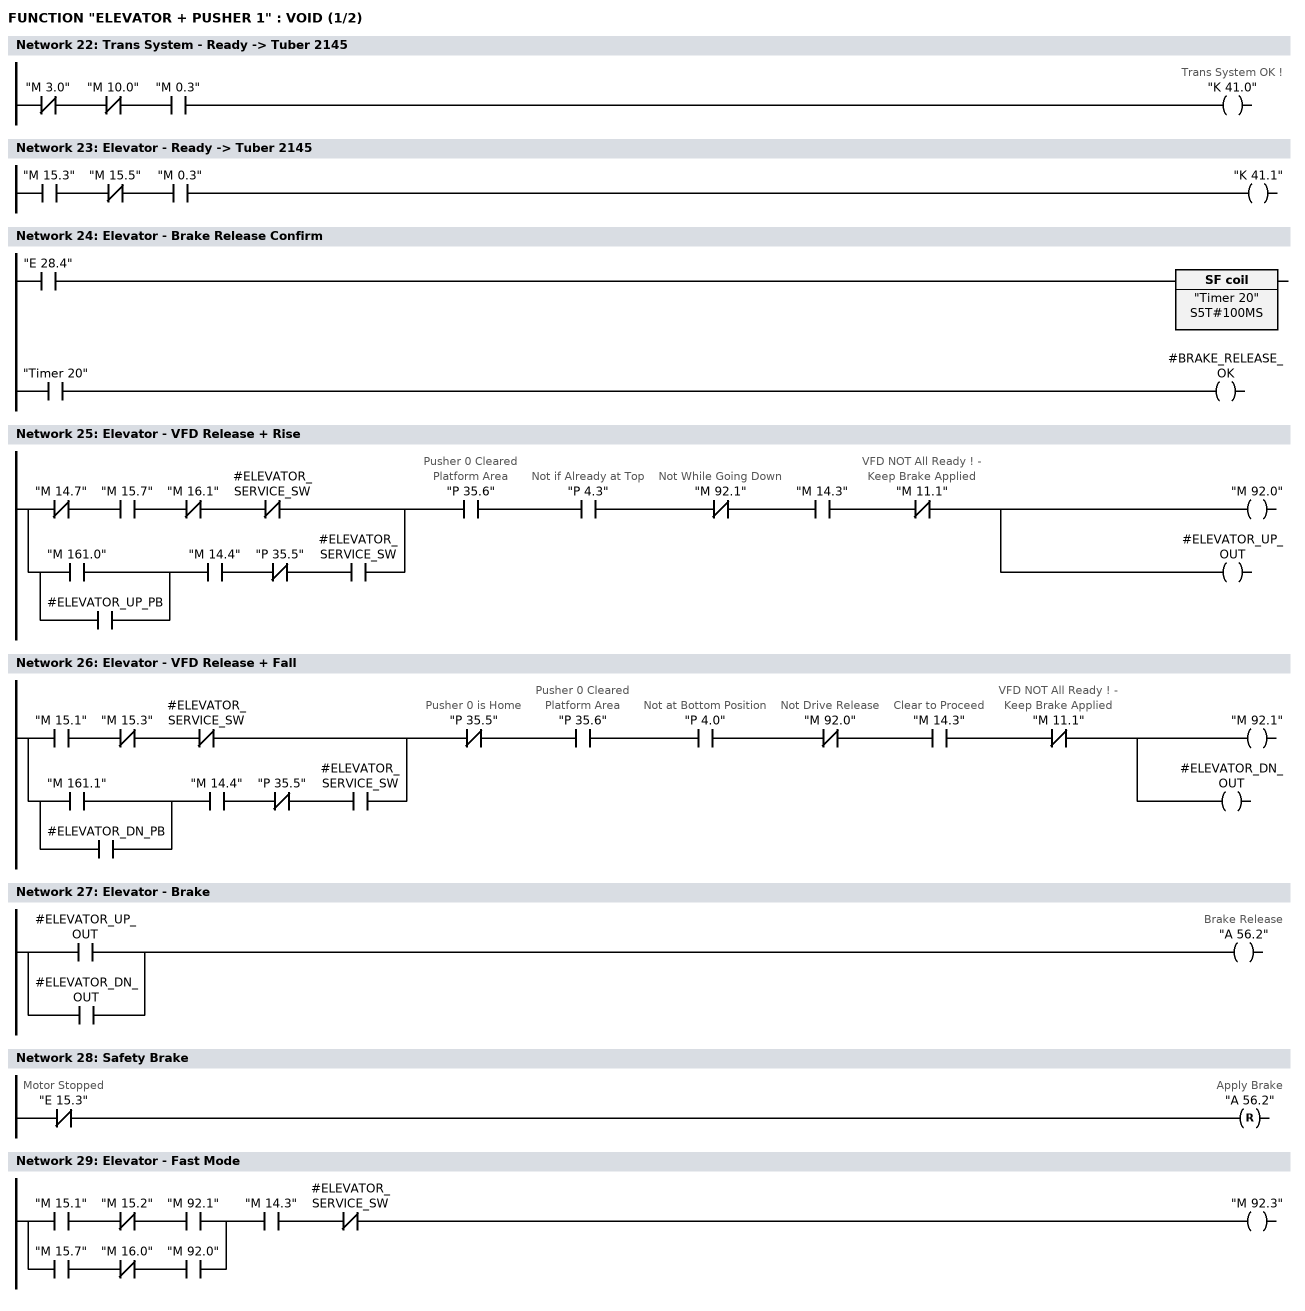

      AN    "M 3.0";
      AN    "M 10.0";
      A     "M 0.3";
      =     "K 41.0"; // Trans System OK !
NETWORK
TITLE =Elevator - Ready -> Tuber 2145

      A     "M 15.3";
      AN    "M 15.5";
      A     "M 0.3";
      =     "K 41.1";
NETWORK
TITLE =Elevator - Brake Release Confirm

      A     "E 28.4";
      L     S5T#100MS;
      SF    "Timer 20";
//;
      A     "Timer 20";
      =     #BRAKE_RELEASE_OK;
NETWORK
TITLE =Elevator - VFD Release + Rise

      A(    ;
      AN    "M 14.7";
      A     "M 15.7";
      AN    "M 16.1";
      AN    #ELEVATOR_SERVICE_SW;
      O     ;
      A(    ;
      O     "M 161.0";
      O     #ELEVATOR_UP_PB;
      )     ;
      A     "M 14.4";
      AN    "P 35.5";
      A     #ELEVATOR_SERVICE_SW;
      )     ;
      A     "P 35.6"; // Pusher 0 Cleared Platform Area
      A     "P 4.3"; // Not if Already at Top
      AN    "M 92.1"; // Not While Going Down
      A     "M 14.3";
      AN    "M 11.1"; // VFD NOT All Ready ! - Keep Brake Applied
      =     "M 92.0";
      =     #ELEVATOR_UP_OUT;
NETWORK
TITLE =Elevator - VFD Release + Fall

      A(    ;
      A     "M 15.1";
      AN    "M 15.3";
      AN    #ELEVATOR_SERVICE_SW;
      O     ;
      A(    ;
      O     "M 161.1";
      O     #ELEVATOR_DN_PB;
      )     ;
      A     "M 14.4";
      AN    "P 35.5";
      A     #ELEVATOR_SERVICE_SW;
      )     ;
      AN    "P 35.5"; // Pusher 0 is Home
      A     "P 35.6"; // Pusher 0 Cleared Platform Area
      A     "P 4.0"; // Not at Bottom Position
      AN    "M 92.0"; // Not Drive Release
      A     "M 14.3"; // Clear to Proceed
      AN    "M 11.1"; // VFD NOT All Ready ! - Keep Brake Applied
      =     "M 92.1";
      =     #ELEVATOR_DN_OUT;
NETWORK
TITLE =Elevator - Brake

      A(    ;
      O     #ELEVATOR_UP_OUT;
      O     #ELEVATOR_DN_OUT;
      )     ;
      =     "A 56.2"; // Brake Release
NETWORK
TITLE =Safety Brake

      AN    "E 15.3"; // Motor Stopped
      R     "A 56.2"; // Apply Brake
NETWORK
TITLE =Elevator - Fast Mode

      A(    ;
      A     "M 15.1";
      AN    "M 15.2";
      A     "M 92.1";
      O     ;
      A     "M 15.7";
      AN    "M 16.0";
      A     "M 92.0";
      )     ;
      A     "M 14.3";
      AN    #ELEVATOR_SERVICE_SW;
      =     "M 92.3";
NETWORK
TITLE =Elevator - Slow
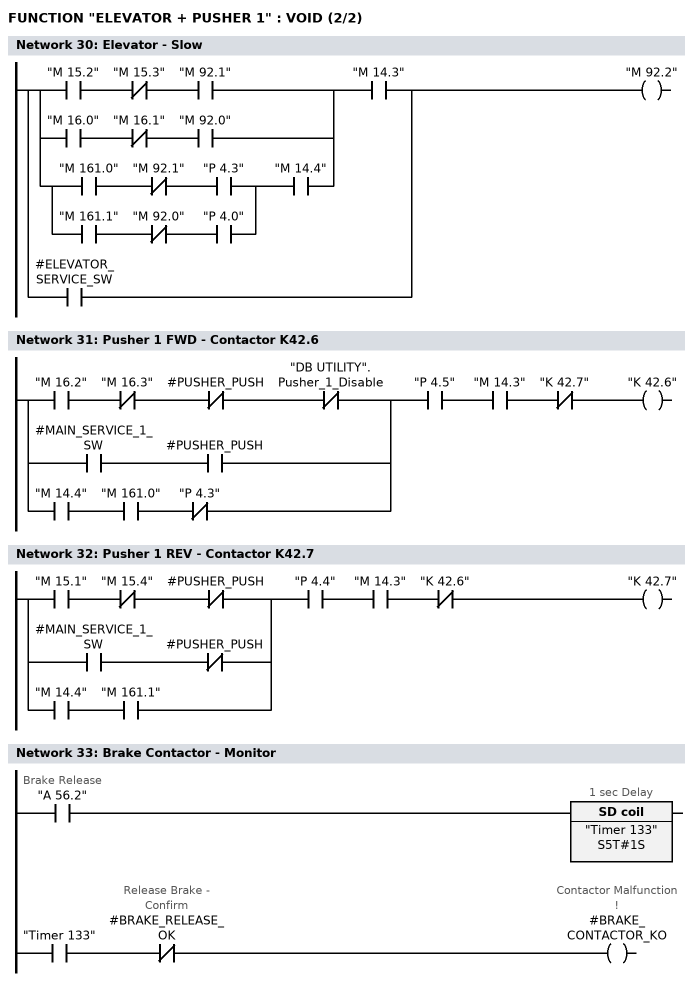

      A(    ;
      A     "M 15.2";
      AN    "M 15.3";
      A     "M 92.1";
      O     ;
      A     "M 16.0";
      AN    "M 16.1";
      A     "M 92.0";
      O     ;
      A(    ;
      A     "M 161.0";
      AN    "M 92.1";
      A     "P 4.3";
      O     ;
      A     "M 161.1";
      AN    "M 92.0";
      A     "P 4.0";
      )     ;
      A     "M 14.4";
      )     ;
      A     "M 14.3";
      O     #ELEVATOR_SERVICE_SW;
      =     "M 92.2";
NETWORK
TITLE =Pusher 1 FWD - Contactor K42.6

      A(    ;
      A     "M 16.2";
      AN    "M 16.3";
      AN    #PUSHER_PUSH;
      AN    "DB UTILITY".Pusher_1_Disable;
      O(    ;
      A     #MAIN_SERVICE_1_SW;
      A     #PUSHER_PUSH;
      )     ;
      O     ;
      A     "M 14.4";
      A     "M 161.0";
      AN    "P 4.3";
      )     ;
      A     "P 4.5";
      A     "M 14.3";
      AN    "K 42.7";
      =     "K 42.6";
NETWORK
TITLE =Pusher 1 REV - Contactor K42.7

      A(    ;
      A     "M 15.1";
      AN    "M 15.4";
      AN    #PUSHER_PUSH;
      O(    ;
      A     #MAIN_SERVICE_1_SW;
      AN    #PUSHER_PUSH;
      )     ;
      O     ;
      A     "M 14.4";
      A     "M 161.1";
      )     ;
      A     "P 4.4";
      A     "M 14.3";
      AN    "K 42.6";
      =     "K 42.7";
NETWORK
TITLE =Brake Contactor - Monitor

      A     "A 56.2"; // Brake Release
      L     S5T#1S; // 1 sec Delay
      SD    "Timer 133";
//;
      A     "Timer 133";
      AN    #BRAKE_RELEASE_OK; // Release Brake - Confirm
      =     #BRAKE_CONTACTOR_KO; // Contactor Malfunction !
NETWORK
TITLE =New Elevator VFD PARKER - Ready

      AN    "E 14.4"; // DRIVE TEST
      O     #BRAKE_CONTACTOR_KO; // Contactor Monitor = Contactor Malfunction !
      JCN   NFLT; // No fault
      S     "M 92.5"; // Set Fault Bit
      JU    OFF; // Turn Off
NETWORK
TITLE =New Elevator VFD with Dynamic Resistor - Go Up

NFLT: A     #ELEVATOR_UP_OUT; // VFD Release Command UP
      A     "M 92.3"; // Fast Speed Command
      AN    "M 92.5"; // Fault Bit
      AN    "M 11.1"; // VFD NOT All Ready !
      JCN   UPLO;
      S     "A 63.0"; // Release Drive - Go Up
      S     "A 63.2"; // Speed 2 / Speed 0.0
//;
      A     #BRAKE_RELEASE_OK; // Release Brake - Confirm
      JCN   END;
      =     "A 63.1"; // Speed 1
      =     "A 63.2"; // Speed 2 + Speed 1 = Fast
      R     "A 63.3"; // L = Forward (Up)
      JU    END;

UPLO: A     #ELEVATOR_UP_OUT; // VFD Release Command UP
      A     "M 92.2"; // Slow Speed Command
      AN    "M 92.5"; // Fault Bit
      AN    "M 11.1"; // VFD NOT All Ready !
      JCN   DNHI;
      S     "A 63.0"; // Release Drive - Go Up
      S     "A 63.2"; // Speed 2 / Speed 0.0
//;
      A     #BRAKE_RELEASE_OK; // Release Brake - Confirm
      JCN   END;
      =     "A 63.1"; // Speed 1
      R     "A 63.2"; // Speed 2 = Off
      R     "A 63.3"; // L = Forward (Up)
      JU    END;
NETWORK
TITLE =New Elevator VFD with Dynamic Resistor - Go Down

DNHI: A     #ELEVATOR_DN_OUT; // VFD Release Command DN
      A     "M 92.3"; // Fast Speed Command
      AN    "M 92.5"; // Fault Bit
      JCN   DNLO;
      S     "A 63.0"; // Release Drive - Go Dn
      S     "A 63.2"; // Speed 2 / Speed 0.0
//;
      A     #BRAKE_RELEASE_OK; // Release Brake - Confirm
      JCN   END;
      =     "A 63.1"; // Speed 1
      =     "A 63.2"; // Speed 2 + Speed 1 = Fast
      =     "A 63.3"; // H = Reverse (Dn)
      JU    END;

DNLO: A     #ELEVATOR_DN_OUT; // VFD Release Command DN
      A     "M 92.2"; // Slow Speed Command
      AN    "M 92.5"; // Fault Bit
      JCN   OFF;
      S     "A 63.0"; // Release Drive - Go Dn
      S     "A 63.2"; // Speed 2 / Speed 0.0
//;
      A     #BRAKE_RELEASE_OK; // Release Brake - Confirm
      JCN   END;
      =     "A 63.1"; // Speed 1
      R     "A 63.2"; // Speed 2 = Off
      =     "A 63.3"; // H = Reverse (Dn)
      JU    END;
NETWORK
TITLE =Drive Off
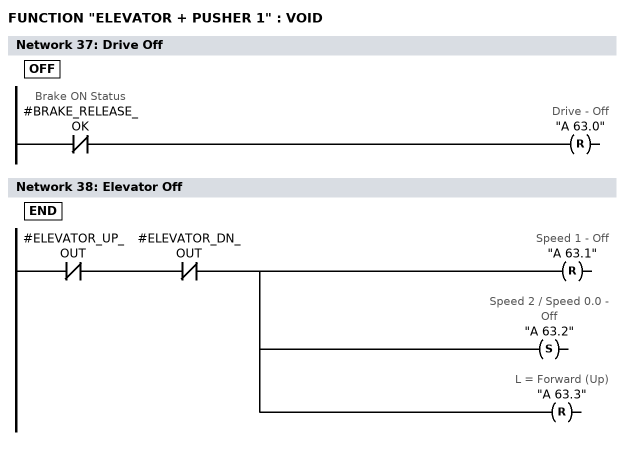

OFF:  AN    #BRAKE_RELEASE_OK; // Brake ON Status
      R     "A 63.0"; // Drive - Off
NETWORK
TITLE =Elevator Off

END:  AN    #ELEVATOR_UP_OUT;
      AN    #ELEVATOR_DN_OUT;
      R     "A 63.1"; // Speed 1 - Off
      S     "A 63.2"; // Speed 2 / Speed 0.0 - Off
      R     "A 63.3"; // L = Forward (Up)
END_FUNCTION

FUNCTION "CONVEYOR 1 - BELT" : VOID
TITLE =Conveyor 1  Pos. 1
//
NAME : POS_3
VERSION : 0.0


VAR_TEMP
  MAIN_SERVICE_1_SW : BOOL ;
  SERVICE_RUN : BOOL ;
  INITIALISATION : BOOL ;
  SENSOR_TEST : BOOL ;
END_VAR
BEGIN
NETWORK
TITLE =Service Test

      A     "HMI_DB".ALL_SERVICE_ENABLE_SW;
      A     "HMI_DB".CONVEYOR_1_SERVICE_SW;
      A     "HMI_DB".SERVICE_SW_1_STATUS;
      =     #MAIN_SERVICE_1_SW;
//;
      A     #MAIN_SERVICE_1_SW;
      O     "M 18.1";
      JNB   CON1;
      A     "HMI_DB".HMI_CONVEYOR_1_TEST_SSW;
      =     #SERVICE_RUN;
      S     "DB UTILITY".Elevator_Disable;
      S     "DB UTILITY".Pusher_1_Disable;
//;
      A     "HMI_DB".SERVICE_INIT_PB;
      =     #INITIALISATION;
//;
      AN    #MAIN_SERVICE_1_SW;
      R     "HMI_DB".HMI_CONVEYOR_1_TEST_SSW;
      R     "DB UTILITY".Elevator_Disable;
      R     "DB UTILITY".Pusher_1_Disable;

CON1: R     #SERVICE_RUN;
      R     #INITIALISATION;
      FP    "FP 158.2";
      =     "M 18.1";
NETWORK
TITLE =Step 2N1 - Power ON
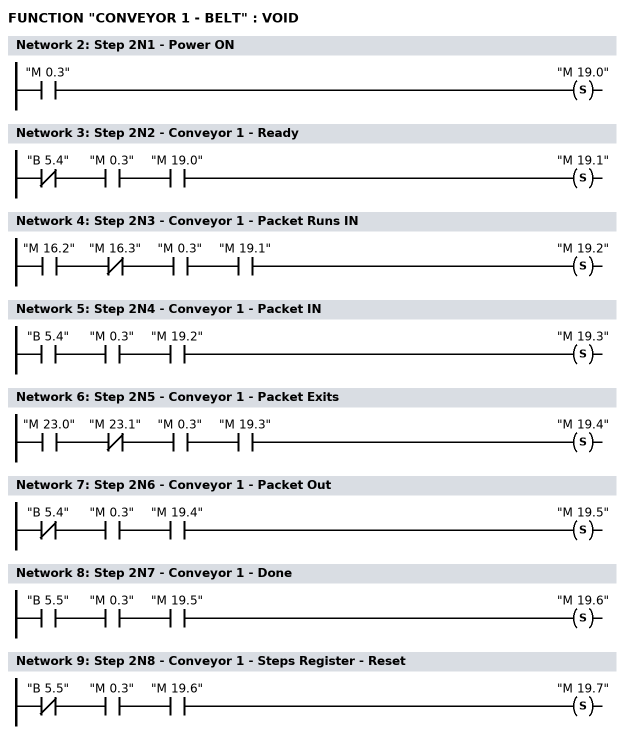

      A     "M 0.3";
      S     "M 19.0";
NETWORK
TITLE =Step 2N2 - Conveyor 1 - Ready

      AN    "B 5.4";
      A     "M 0.3";
      A     "M 19.0";
      S     "M 19.1";
NETWORK
TITLE =Step 2N3 - Conveyor 1 - Packet Runs IN

      A     "M 16.2";
      AN    "M 16.3";
      A     "M 0.3";
      A     "M 19.1";
      S     "M 19.2";
NETWORK
TITLE =Step 2N4 - Conveyor 1 - Packet IN

      A     "B 5.4";
      A     "M 0.3";
      A     "M 19.2";
      S     "M 19.3";
NETWORK
TITLE =Step 2N5 - Conveyor 1 - Packet Exits

      A     "M 23.0";
      AN    "M 23.1";
      A     "M 0.3";
      A     "M 19.3";
      S     "M 19.4";
NETWORK
TITLE =Step 2N6 - Conveyor 1 - Packet Out

      AN    "B 5.4";
      A     "M 0.3";
      A     "M 19.4";
      S     "M 19.5";
NETWORK
TITLE =Step 2N7 - Conveyor 1 - Done

      A     "B 5.5";
      A     "M 0.3";
      A     "M 19.5";
      S     "M 19.6";
NETWORK
TITLE =Step 2N8 - Conveyor 1 - Steps Register - Reset

      AN    "B 5.5";
      A     "M 0.3";
      A     "M 19.6";
      S     "M 19.7";
NETWORK
TITLE =Conveyor 1 - Steps Register - Reset

      A(    ;
      O     "M 19.7";
      O     "DB UTILITY".T19_DN;
      O     #INITIALISATION;
      O     "DB UTILITY".Conveyor_1_Disable;
      )     ;
      A     "M 0.3";
      JNB   INIT;
      L     W#16#0;
      T     "MW 19";

INIT: CLR   ;
NETWORK
TITLE =Soft Timer 19 Reset

      A     "M 19.2";
      AN    "M 19.3";
      A     "M 0.3";
      JCN   R191;
      JU    E191;

R191: L     L#0;
      T     "DB UTILITY".T19_ET;
      R     "DB UTILITY".T19_DN;

E191: NOP   0;

NETWORK
TITLE =Soft Timer 19 Add

      A     "M 19.2";
      AN    "M 19.3";
      A     "M 0.3";
      AN    "DB UTILITY".Freeze_Sequence_1;
      AN    "DB UTILITY".T19_DN;
      JCN   E192;

      L     "DB UTILITY".T19_ET;
      L     "DB UTILITY".Scan_Cycle_Previous;
      ITD   ;
      +D    ;
      T     "DB UTILITY".T19_ET;

E192: NOP   0;

NETWORK
TITLE =Soft Timer 19 Done 10s
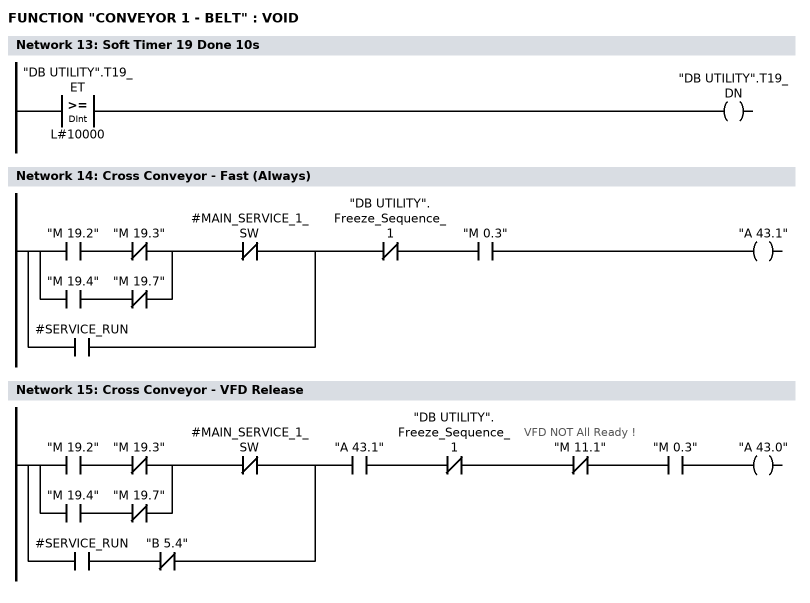

      L     "DB UTILITY".T19_ET;
      L     L#10000;
      >=D   ;
      =     "DB UTILITY".T19_DN;
NETWORK
TITLE =Cross Conveyor - Fast (Always)

      A(    ;
      A     "M 19.2";
      AN    "M 19.3";
      O     ;
      A     "M 19.4";
      AN    "M 19.7";
      )     ;
      AN    #MAIN_SERVICE_1_SW;
      O     #SERVICE_RUN;
      AN    "DB UTILITY".Freeze_Sequence_1;
      A     "M 0.3";
      =     "A 43.1";

NETWORK
TITLE =Cross Conveyor - VFD Release

      A(    ;
      A     "M 19.2";
      AN    "M 19.3";
      O     ;
      A     "M 19.4";
      AN    "M 19.7";
      )     ;
      AN    #MAIN_SERVICE_1_SW;
      O(    ;
      A     #SERVICE_RUN;
      AN    "B 5.4";
      )     ;
      A     "A 43.1";
      AN    "DB UTILITY".Freeze_Sequence_1;
      AN    "M 11.1"; // VFD NOT All Ready !
      A     "M 0.3";
      =     "A 43.0";
NETWORK
TITLE =Any Conveyors Packet mS Test

//    A     "B 10.7"
//    A     "A 48.6"


      A     "B 10.6";
      A     "A 48.3";






      =     #SENSOR_TEST;
//;
      A     #SENSOR_TEST;
      FP    "FP 147.7";
      JNB   NRST;
      L     0;
      T     "COLLATORS DB".Any_Conveyors_mS;

NRST: A     #SENSOR_TEST;
      JNB   NCNT;
      L     "COLLATORS DB".Any_Conveyors_mS;
      L     "DB UTILITY".Scan_Cycle_Previous;
      ITD   ;
      +D    ;
      T     "COLLATORS DB".Any_Conveyors_mS;

NCNT: CLR   ;

END_FUNCTION

FUNCTION "CONVEYOR 2 - ANGLE B+R" : VOID
TITLE =Angle Conveyor 2  Pos. 4
NAME : POS_4
VERSION : 0.0


VAR_TEMP
  MAIN_SERVICE_1_SW : BOOL ;
  SERVICE_BELT_RUN : BOOL ;
  SERVICE_ROLLER_LIFT : BOOL ;
  SERVICE_ROLLER_RUN : BOOL ;
  INITIALISATION : BOOL ;
  PACKET_MEASURE_FLAG : BOOL ;
END_VAR
BEGIN
NETWORK
TITLE =Service Test

      A     "HMI_DB".ALL_SERVICE_ENABLE_SW;
      A     "HMI_DB".CONVEYOR_2_SERVICE_SW;
      A     "HMI_DB".SERVICE_SW_1_STATUS;
      =     #MAIN_SERVICE_1_SW;
//;
      A     #MAIN_SERVICE_1_SW;
      O     "M 22.1";
      JNB   CON2;
      A     "HMI_DB".HMI_CONVEYOR_2B_TEST_SSW;
      =     #SERVICE_BELT_RUN;
      S     "DB UTILITY".Conveyor_1_Disable;
//;
      A     "HMI_DB".HMI_CONVEYOR_2L_TEST_SSW;
      =     #SERVICE_ROLLER_LIFT;
      S     "DB UTILITY".Conveyor_1_Disable;
//;
      A     "HMI_DB".HMI_CONVEYOR_2R_TEST_SSW;
      =     #SERVICE_ROLLER_RUN;
      S     "DB UTILITY".Conveyor_1_Disable;
//;
      A     "HMI_DB".SERVICE_INIT_PB;
      =     #INITIALISATION;
//;
      AN    #MAIN_SERVICE_1_SW;
      R     "HMI_DB".HMI_CONVEYOR_2B_TEST_SSW;
      R     "HMI_DB".HMI_CONVEYOR_2L_TEST_SSW;
      R     "HMI_DB".HMI_CONVEYOR_2R_TEST_SSW;
      R     "DB UTILITY".Conveyor_1_Disable;

CON2: R     #SERVICE_BELT_RUN;
      R     #SERVICE_ROLLER_LIFT;
      R     #SERVICE_ROLLER_RUN;
      R     #INITIALISATION;
      FP    "FP 158.3";
      =     "M 22.1";

NETWORK
TITLE =Angle Conveyor - Fault / Ready
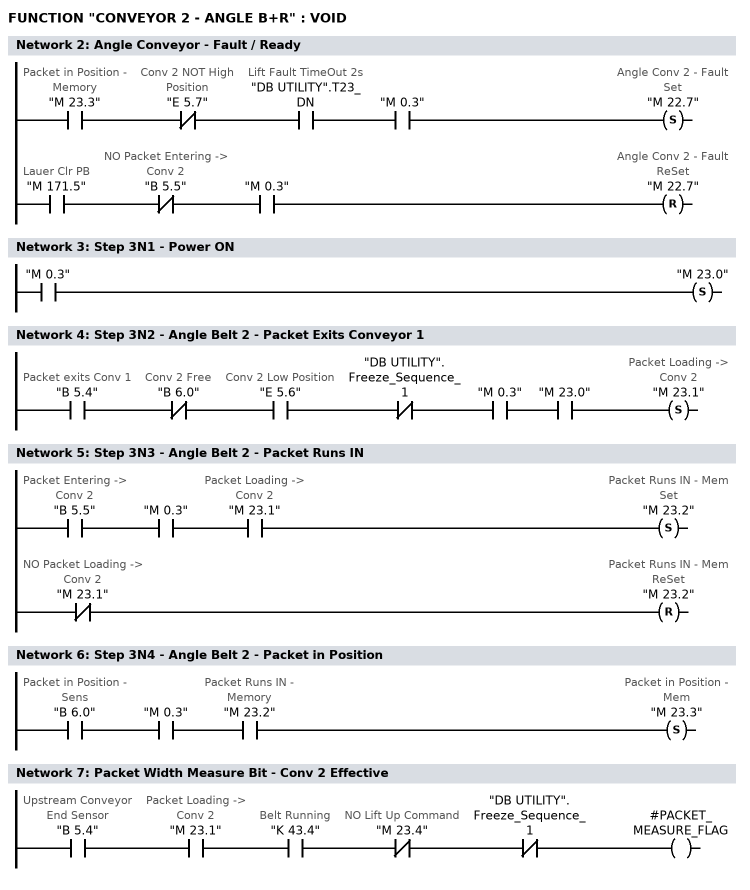

      A     "M 23.3"; // Packet in Position - Memory
      AN    "E 5.7"; // Conv 2 NOT High Position
      A     "DB UTILITY".T23_DN; // Lift Fault TimeOut 2s
      A     "M 0.3";
      S     "M 22.7"; // Angle Conv 2 - Fault Set
//;
      A     "M 171.5"; // Lauer Clr PB
      AN    "B 5.5"; // NO Packet Entering -> Conv 2
      A     "M 0.3";
      R     "M 22.7"; // Angle Conv 2 - Fault ReSet

NETWORK
TITLE =Step 3N1 - Power ON

      A     "M 0.3";
      S     "M 23.0";

NETWORK
TITLE =Step 3N2 - Angle Belt 2 - Packet Exits Conveyor 1

      A     "B 5.4"; // Packet exits Conv 1
      AN    "B 6.0"; // Conv 2 Free
      A     "E 5.6"; // Conv 2 Low Position
      AN    "DB UTILITY".Freeze_Sequence_1;
      A     "M 0.3";
      A     "M 23.0";
      S     "M 23.1"; // Packet Loading -> Conv 2
NETWORK
TITLE =Step 3N3 - Angle Belt 2 - Packet Runs IN

      A     "B 5.5"; // Packet Entering -> Conv 2
      A     "M 0.3";
      A     "M 23.1"; // Packet Loading -> Conv 2
      S     "M 23.2"; // Packet Runs IN - Mem Set
//;
      ON    "M 23.1"; // NO Packet Loading -> Conv 2
      R     "M 23.2"; // Packet Runs IN - Mem ReSet

NETWORK
TITLE =Step 3N4 - Angle Belt 2 - Packet in Position

      A     "B 6.0"; // Packet in Position - Sens
      A     "M 0.3";
      A     "M 23.2"; // Packet Runs IN - Memory
      S     "M 23.3"; // Packet in Position - Mem
NETWORK
TITLE =Packet Width Measure Bit - Conv 2 Effective

      A     "B 5.4"; // Upstream Conveyor End Sensor
      A     "M 23.1"; // Packet Loading -> Conv 2
      A     "K 43.4"; // Belt Running
      AN    "M 23.4"; // NO Lift Up Command
      AN    "DB UTILITY".Freeze_Sequence_1;
      =     #PACKET_MEASURE_FLAG;

NETWORK
TITLE =Packet Width Time Reset - Freeze Safe

      A     "M 23.1"; // Packet Loading -> Conv 2
      O     "DB UTILITY".Freeze_Sequence_1;
      JC    NRS1;

      L     L#0;
      T     "MD 260"; // Width [mS]

NRS1: NOP   0;
NETWORK
TITLE =Packet Width Time Count Up From Sensor "B 5.4"

      A     #PACKET_MEASURE_FLAG;
      JCN   NMES;

      L     "MD 260"; // Width [mS]
      L     "DB UTILITY".Scan_Cycle_Previous;
      ITD   ;
      +D    ;
      T     "MD 260"; // Width [mS]

NMES: NOP   0;
NETWORK
TITLE =Middle Travel Time Reset - Freeze Safe

      A     "M 23.3"; // Packet in Position - Mem
      O     "DB UTILITY".Freeze_Sequence_1;
      JC    NRS2;

      L     L#0;
      T     "MD 264"; // Half Width [mS] - Zeroed

NRS2: NOP   0;
NETWORK
TITLE =Middle Travel Time Count Up From B 6.0

      ON    "M 23.3"; // NO Packet in Position - Mem
      O     "M 23.4"; // Lift Up Command
      ON    "K 43.4"; // Belt Stopped
      ON    "M 0.3"; // No Power
      AN    "DB UTILITY".Freeze_Sequence_1;
      JC    NCNT;

      L     "MD 264"; // Half Width [mS]
      L     "DB UTILITY".Scan_Cycle_Previous;
      ITD   ;
      +D    ;
      T     "MD 264"; // Half Width [mS] - Add

NCNT: NOP   0;
NETWORK
TITLE =Middle Travel Time Clamp Zero

      L     "MD 264"; // Half Width [mS]
      L     L#0;
      >=D   ;
      JC    NMID;

      L     L#0;
      T     "MD 264"; // Half Width [mS] - Reset

NMID: NOP   0;
NETWORK
TITLE =Soft Timer 23 Reset - Lift Fault TimeOut 2s + Freeze Option

      A     "M 23.3"; // Packet in Position - Memory
      AN    "M 23.4"; // NO Lift Up Command
      A     "M 0.3";
      JCN   R231;
      JU    E231;

R231: L     L#0;
      T     "DB UTILITY".T23_ET;
      R     "DB UTILITY".T23_DN;

E231: NOP   0;

NETWORK
TITLE =Soft Timer 23 Add

      A     "M 23.3"; // Packet in Position - Memory
      AN    "M 23.4"; // NO Lift Up Command
      A     "M 0.3";
      AN    "DB UTILITY".Freeze_Sequence_1; // Sequence Freezer Bit
      AN    "DB UTILITY".T23_DN;
      JCN   E232;

      L     "DB UTILITY".T23_ET;
      L     "DB UTILITY".Scan_Cycle_Previous;
      ITD   ;
      +D    ;
      T     "DB UTILITY".T23_ET;

E232: NOP   0;

NETWORK
TITLE =Soft Timer 23 Done 2s

      L     "DB UTILITY".T23_ET;
      L     L#2500; // [mS]
      >=D   ;
      =     "DB UTILITY".T23_DN;
NETWORK
TITLE =Soft Timer 24 Reset - Belt TimeOut 8s + Freeze Option

      A     "M 23.1";
      AN    "M 23.3";
      A     "K 43.4";
      A     "M 0.3";
      JCN   R241;
      JU    E241;

R241: L     L#0;
      T     "DB UTILITY".T24_ET;
      R     "DB UTILITY".T24_DN;

E241: NOP   0;

NETWORK
TITLE =Soft Timer 24 Add

      A     "M 23.1";
      AN    "M 23.3";
      A     "K 43.4";
      A     "M 0.3";
      AN    "DB UTILITY".Freeze_Sequence_1;
      AN    "DB UTILITY".T24_DN;
      JCN   E242;

      L     "DB UTILITY".T24_ET;
      L     "DB UTILITY".Scan_Cycle_Previous;
      ITD   ;
      +D    ;
      T     "DB UTILITY".T24_ET;

E242: NOP   0;

NETWORK
TITLE =Soft Timer 24 Done 8s

      L     "DB UTILITY".T24_ET;
      L     L#8000;
      >=D   ;
      =     "DB UTILITY".T24_DN;
      S     "M 24.4";
NETWORK
TITLE =Step 3N5 - Angle Belt - Lift ("MD 264" to Center the Packet)

      A(    ;
      A(    ;
      L     "MD 264";
      L     L#2;
      *D    ;
      L     "MD 260";
      >=D   ;
      )     ;
      AN    #PACKET_MEASURE_FLAG;
      AN    "B 5.5";
      O     "DB UTILITY".T23_DN;
      )     ;
      A     "M 0.3";
      A     "M 23.3";
      S     "M 23.4";
NETWORK
TITLE =Step 3N6 - Angle Rollers - Up
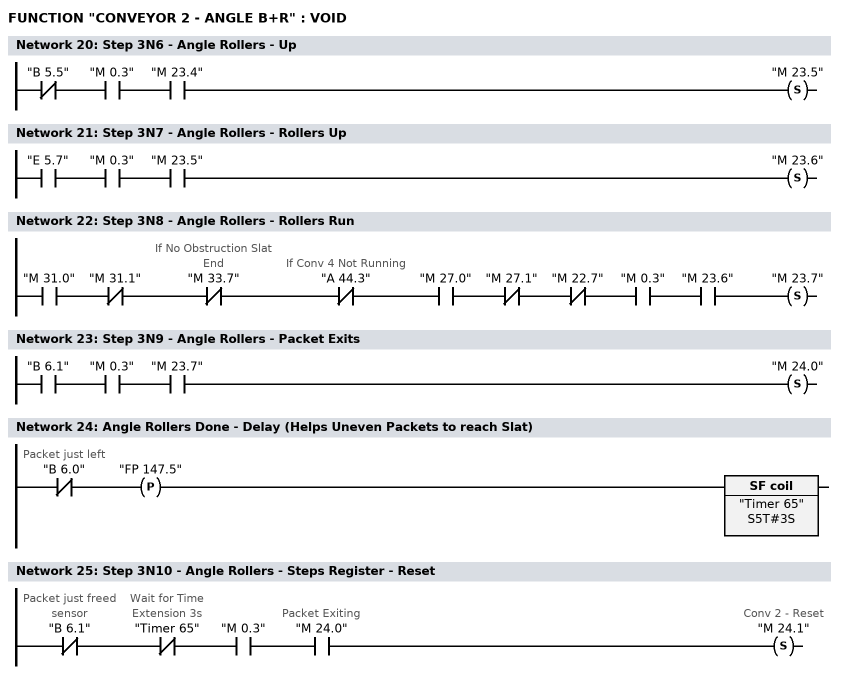

      AN    "B 5.5";
      A     "M 0.3";
      A     "M 23.4";
      S     "M 23.5";

NETWORK
TITLE =Step 3N7 - Angle Rollers - Rollers Up

      A     "E 5.7";
      A     "M 0.3";
      A     "M 23.5";
      S     "M 23.6";

NETWORK
TITLE =Step 3N8 - Angle Rollers - Rollers Run

      A     "M 31.0";
      AN    "M 31.1";
      AN    "M 33.7"; // If No Obstruction Slat End
      AN    "A 44.3"; // If Conv 4 Not Running
      A     "M 27.0";
      AN    "M 27.1";
      AN    "M 22.7";
      A     "M 0.3";
      A     "M 23.6";
      S     "M 23.7";

NETWORK
TITLE =Step 3N9 - Angle Rollers - Packet Exits

      A     "B 6.1";
      A     "M 0.3";
      A     "M 23.7";
      S     "M 24.0";

NETWORK
TITLE =Angle Rollers Done - Delay (Helps Uneven Packets to reach Slat)

      AN    "B 6.0"; // Packet just left
      FP    "FP 147.5";
      L     S5T#3S;
      SF    "Timer 65"; // Time Extension 3s
NETWORK
TITLE =Step 3N10 - Angle Rollers - Steps Register - Reset

      AN    "B 6.1"; // Packet just freed sensor
      AN    "Timer 65"; // Wait for Time Extension 3s
      A     "M 0.3";
      A     "M 24.0"; // Packet Exiting
      S     "M 24.1"; // Conv 2 - Reset
NETWORK
TITLE =Conveyor 2 - Steps Register - Reset

      A(    ;
      O     "M 24.1";
      O     "DB UTILITY".T24_DN;
      O     "DB UTILITY".T25_DN;
      O     #INITIALISATION;
      O     "DB UTILITY".Conveyor_1_Disable;
      )     ;
      A     "M 0.3";
      JC    M001;
      JU    M002;

M001: L     W#16#0;
      T     "MW 23";

M002: NOP   0;
NETWORK
TITLE =Soft Timer 25 Reset - Roller TimeOut 8s + Freeze Option

      A     "M 23.7";
      AN    "M 24.1";
      A     "M 0.3";
      JCN   R251;
      JU    E251;

R251: L     L#0;
      T     "DB UTILITY".T25_ET;
      R     "DB UTILITY".T25_DN;

E251: NOP   0;

NETWORK
TITLE =Soft Timer 25 Add

      A     "M 23.7";
      AN    "M 24.1";
      A     "M 0.3";
      AN    "DB UTILITY".Freeze_Sequence_2;
      AN    "DB UTILITY".T25_DN;
      JCN   E252;

      L     "DB UTILITY".T25_ET;
      L     "DB UTILITY".Scan_Cycle_Previous;
      ITD   ;
      +D    ;
      T     "DB UTILITY".T25_ET;

E252: NOP   0;

NETWORK
TITLE =Soft Timer 25 Done 8s

      L     "DB UTILITY".T25_ET;
      L     L#8000;
      >=D   ;
      =     "DB UTILITY".T25_DN;
NETWORK
TITLE =Angle Conveyor Belt - Run

      A     "M 23.1";
      AN    "M 23.4";
      AN    #MAIN_SERVICE_1_SW;
      O(    ;
      A     #SERVICE_BELT_RUN;
      A(    ;
      A     "B 6.0";
      L     S5T#200MS;
      SD    "Timer 21";
//;
      AN    "Timer 21";
      )     ;
      )     ;
      AN    "M 22.7";
      AN    "DB UTILITY".Freeze_Sequence_1;
      AN    "M 11.1"; // VFD NOT All Ready !
      A     "M 0.3";
      =     "K 43.4";

NETWORK
TITLE =Angle Conveyor Rollers - Run
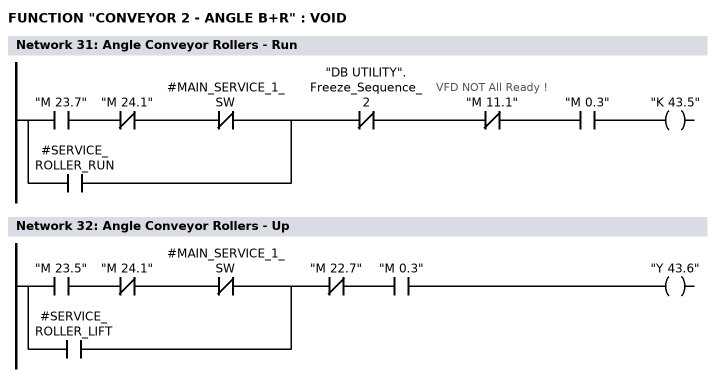

      A     "M 23.7";
      AN    "M 24.1";
      AN    #MAIN_SERVICE_1_SW;
      O     #SERVICE_ROLLER_RUN;
      AN    "DB UTILITY".Freeze_Sequence_2;
      AN    "M 11.1"; // VFD NOT All Ready !
      A     "M 0.3";
      =     "K 43.5";

NETWORK
TITLE =Angle Conveyor Rollers - Up

      A     "M 23.5";
      AN    "M 24.1";
      AN    #MAIN_SERVICE_1_SW;
      O     #SERVICE_ROLLER_LIFT;
      AN    "M 22.7";
      A     "M 0.3";
      =     "Y 43.6";
END_FUNCTION

FUNCTION "CONVEYOR 3 - SLAT" : VOID
TITLE =Slat Conveyor 3  Pos.5
NAME : POS_5
VERSION : 0.0


VAR_TEMP
  MAIN_SERVICE_1_SW : BOOL ;
  SERVICE_RUN : BOOL ;
  INITIALISATION : BOOL ;
END_VAR
BEGIN
NETWORK
TITLE =Service Test

      A     "HMI_DB".ALL_SERVICE_ENABLE_SW;
      A     "HMI_DB".CONVEYOR_3_SERVICE_SW;
      A     "HMI_DB".SERVICE_SW_1_STATUS;
      =     #MAIN_SERVICE_1_SW;
//;
      A     #MAIN_SERVICE_1_SW;
      O     M     26.3;
      JNB   CON3;
      A     "HMI_DB".HMI_CONVEYOR_3_TEST_SSW;
      =     #SERVICE_RUN;
      S     "DB UTILITY".Conveyor_2_Disable;
//;
      AN    #MAIN_SERVICE_1_SW;
      R     "HMI_DB".HMI_CONVEYOR_3_TEST_SSW;
      R     "DB UTILITY".Conveyor_2_Disable;
//;
      A     "HMI_DB".SERVICE_INIT_PB;
      A     #MAIN_SERVICE_1_SW;
      =     #INITIALISATION;

CON3: R     #SERVICE_RUN;
      FP    "FP 227.0";
      =     M     26.3;
NETWORK
TITLE =Packet Length Measurements [mm] - While Collating

      A     "B 6.2"; // C3 InFeed Sens - New Packet
      FP    "FP 227.1";
      A     "A 44.0";
      JC    PRNT;
      JU    RPRT;

PRNT: L     "FM350 DB".ACT_CNTV0;
      T     "HOUSE_KEEPING DB".C3_Encoder_READ_Mem;

RPRT: AN    "B 6.2"; // C3 InFeed Sens - New Packet End
      FP    "FP 227.2";
      JCN   NTKE;

      L     "FM350 DB".ACT_CNTV0;
      L     "HOUSE_KEEPING DB".C3_Encoder_READ_Mem;
      -I    ;
      T     "HOUSE_KEEPING DB".C3_Packet_Length_ep;
      DTR   ;
//;
      L     1.300000e+00; //  Encoder Wheel 900mm / 600 PPR  [mm/pulse]
      *R    ;
      RND   ;
      T     "HOUSE_KEEPING DB".C3_Packet_Length_mm;

NTKE: NOP   0;
NETWORK
TITLE =Slat Conveyor 3 - Packets / Conveyor Length - Calculation

      A     "M 27.1";
      FP    "FP 227.3";
      JNB   M271;
      L     "COLLATORS DB".Conveyor_Length_C3;
      ITD   ;
      DTR   ;
      L     5.000000e+00;
      /R    ;
      RND   ;
      T     "COLLATORS DB".Press_Length_C3;
      T     "MW 212";

M271: NOP   0;
NETWORK
TITLE =Slat Conveyor 3 - Surface Length Manager (PulseUnit)

      A     "M 27.1";
      O     "M 26.6";
      S     "M 166.0";
//;
      A     "M 166.0";
      O(    ;
      AN    "M 10.0";
      FP    "FP 227.4";
      )     ;
      =     "FM350 DB".CONTROL_SIGNALS.SW_GATE0; // C3 Surface Count
//;



////////////////////////////////////////


      A     "M 166.0"; // Start Count (100mS Pulse)
      A(    ;
      L     "FM350 DB".ACT_CNTV0; // C3 Surface Count
      L     "MW 212";
      >=I   ;
      )     ;
      A     "M 0.3";
      JCN   R291;
      JU    E291;

R291: L     L#0;
      T     "DB UTILITY".T27_ET;
      R     "DB UTILITY".T27_DN;

E291: NOP   0;

NETWORK
TITLE =Soft Timer 27 Add - FM350 needs a 100mS Pulse !

      A     "M 166.0";
      A(    ;
      L     "FM350 DB".ACT_CNTV0; // C3 Surface Count
      L     "MW 212";
      >=I   ;
      )     ;
      A     "M 0.3";
      AN    "DB UTILITY".Freeze_Sequence_2;
      AN    "DB UTILITY".T27_DN;
      JCN   E292;

      L     "DB UTILITY".T27_ET;
      L     "DB UTILITY".Scan_Cycle_Previous;
      ITD   ;
      +D    ;
      T     "DB UTILITY".T27_ET;

E292: NOP   0;

NETWORK
TITLE =Soft Timer 27 Done 100mS  // Start Count (100mS Pulse)
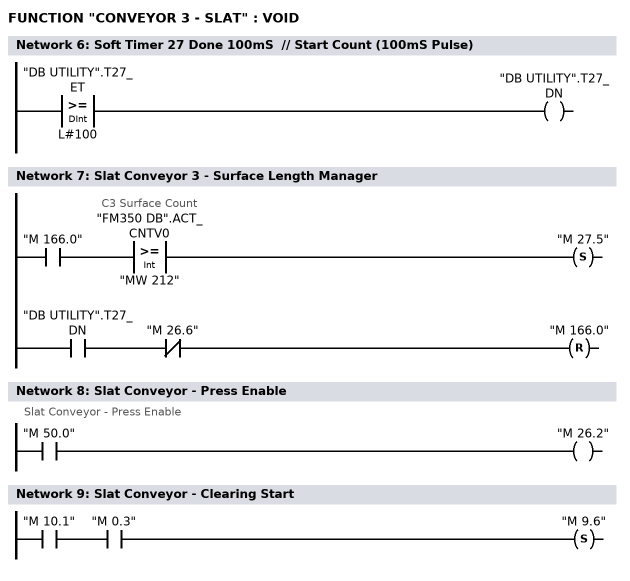

      L     "DB UTILITY".T27_ET;
      L     L#100;
      >=D   ;
      =     "DB UTILITY".T27_DN;

NETWORK
TITLE =Slat Conveyor 3 - Surface Length Manager

      A     "M 166.0";
      A(    ;
      L     "FM350 DB".ACT_CNTV0; // C3 Surface Count
      L     "MW 212";
      >=I   ;
      )     ;
      S     "M 27.5";
//;
      A     "DB UTILITY".T27_DN;
      AN    "M 26.6";
      R     "M 166.0";




////////////////////////////////////////




NETWORK
TITLE =Slat Conveyor - Press Enable
//Slat Conveyor - Press Enable
      A     "M 50.0";
      =     "M 26.2";
NETWORK
TITLE =Slat Conveyor - Clearing Start

      A     "M 10.1";
      A     "M 0.3";
      S     "M 9.6";
NETWORK
TITLE =Slat Conveyor - Clearing
//Counting 9K Pulses Should Suffice !
      A     "M 10.1";
      AN    "M 10.2";
      AN    "A 44.0";
      S     "M 26.6";
//;
      A     "M 26.6";
      JNB   M266;
      A(    ;
      L     "FM350 DB".ACT_CNTV0; // C3 Surface Count
      L     10000;
      >I    ;
      )     ;
      =     "M 26.7";

M266: NOP   0;

      A     "M 26.7";
      ON    "M 10.0";
      R     "M 26.6";
NETWORK
TITLE =Slat Conveyor Steps
//Slat Conveyor Steps


NETWORK
TITLE =Step 4N1 - Power ON
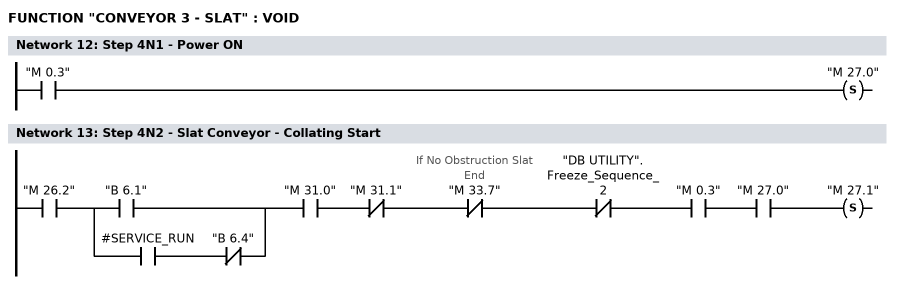

      A     "M 0.3";
      S     "M 27.0";
NETWORK
TITLE =Step 4N2 - Slat Conveyor - Collating Start

      A     "M 26.2";
      A(    ;
      O     "B 6.1";
      O(    ;
      A     #SERVICE_RUN;
      AN    "B 6.4";
      )     ;
      )     ;
      A     "M 31.0";
      AN    "M 31.1";
      AN    "M 33.7"; // If No Obstruction Slat End
      AN    "DB UTILITY".Freeze_Sequence_2;
      A     "M 0.3";
      A     "M 27.0";
      S     "M 27.1";



////////////////////////////////////////



NETWORK
TITLE =Soft Timer 28 Reset - Collating TimeOut + Freeze Option

      A     "M 27.1";
      AN    "M 27.4";
      A     "M 0.3";
      JCN   R271;
      JU    E271;

R271: L     L#0;
      T     "DB UTILITY".T28_ET;
      R     "DB UTILITY".T28_DN;

E271: NOP   0;

NETWORK
TITLE =Soft Timer 28 Add

      A     "M 27.1";
      AN    "M 27.4";
      A     "M 0.3";
      AN    "DB UTILITY".Freeze_Sequence_2;
      AN    "DB UTILITY".T28_DN;
      JCN   E272;

      L     "DB UTILITY".T28_ET;
      L     "DB UTILITY".Scan_Cycle_Previous;
      ITD   ;
      +D    ;
      T     "DB UTILITY".T28_ET;

E272: NOP   0;

NETWORK
TITLE =Soft Timer 27 Done 11s
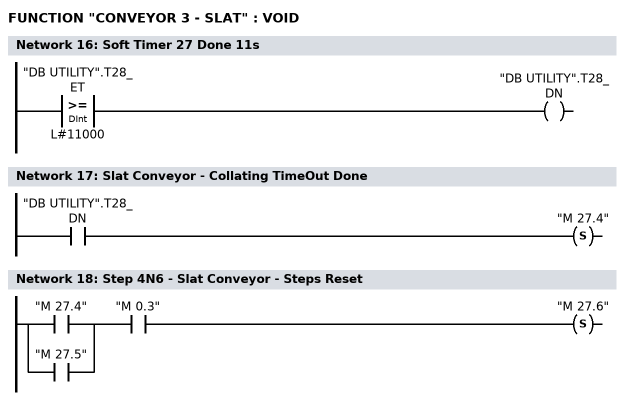

      L     "DB UTILITY".T28_ET;
      L     L#11000;
      >=D   ;
      =     "DB UTILITY".T28_DN;

NETWORK
TITLE =Slat Conveyor - Collating TimeOut Done

      A     "DB UTILITY".T28_DN;
      S     "M 27.4";



////////////////////////////////////////




NETWORK
TITLE =Step 4N6 - Slat Conveyor - Steps Reset

      O     "M 27.4";
      O     "M 27.5";
      A     "M 0.3";
      S     "M 27.6";
NETWORK
TITLE =Slat Conveyor - Steps Register - Reset

      A(    ;
      O     "M 27.6";
      O     #INITIALISATION;
      O     "DB UTILITY".Conveyor_3_Disable;
      )     ;
      A     "M 0.3";
      JC    M001;
      JU    M002;

M001: L     W#16#0;
      T     "MB 27";
      R     "M 26.7";

M002: NOP   0;
NETWORK
TITLE =Slat Conveyor - VFD Release

      A(    ;
      O     "M 27.1";
      O     "M 26.6";
      )     ;
      AN(   ;
      A     "M 26.6";
      A     "M 31.5";
      )     ;
      AN    "DB UTILITY".Freeze_Sequence_2;
      AN    "M 11.1"; // VFD NOT All Ready !
      A     "M 0.3";
      =     "A 44.0";
      =     "A 44.1";
END_FUNCTION

FUNCTION "CONVEYOR 4 - COLLATOR" : VOID
TITLE =Collator Conveyor 4  Pos.6
//Collator Conveyor 4 - Is On Both Service Pages 1 & 2
NAME : POS_6
VERSION : 0.0


VAR_TEMP
  MAIN_SERVICE_1_2_SW : BOOL ;	//Collator Conveyor 4 - On Service 1 & 2
  SERVICE_RUN : BOOL ;
  INITIALISATION : BOOL ;
  COUNTER_TRIGGER : BOOL ;
  PACKET_LENGTH_4 : WORD ;	//Collator Conveyor 4 - Packet Length
  W_TUBE_mm : WORD ;
  W_TUBE_PERCENT : WORD ;	//Tube 5 % Value
  R_TUBE_PERCENT : REAL ;	//Tube 5 % Value
  R_TUBE_mm : REAL ;
END_VAR
BEGIN
NETWORK
TITLE =Conveyor 4 - Service

      A     "HMI_DB".ALL_SERVICE_ENABLE_SW;
      A     "HMI_DB".CONVEYOR_4_SERVICE_SW;
      A(    ;
      O     "HMI_DB".SERVICE_SW_1_STATUS;
      O     "HMI_DB".SERVICE_SW_2_STATUS;
      )     ;
      =     "HMI_DB".SERVICE_SW_1_2_STATUS;
      =     #MAIN_SERVICE_1_2_SW;
//;
      A     #MAIN_SERVICE_1_2_SW;
      O     "M 26.1";
      JNB   CON4;
      A     "HMI_DB".HMI_CONVEYOR_4_TEST_SSW;
      =     #SERVICE_RUN;
      S     "DB UTILITY".Conveyor_3_Disable;
//;
      A     "HMI_DB".SERVICE_INIT_PB;
      A     #MAIN_SERVICE_1_2_SW;
      =     #INITIALISATION;
//;
      AN    #MAIN_SERVICE_1_2_SW;
      R     "HMI_DB".HMI_CONVEYOR_4_TEST_SSW;
      R     "DB UTILITY".Conveyor_3_Disable;

CON4: R     #SERVICE_RUN;
      R     #INITIALISATION;
      FP    "FP 158.4";
      =     "M 26.1";
NETWORK
TITLE =Soft Timer 90 Reset Conveyor 4 - Encoder has Stop L - Timer  500

      AN    "E 6.6";
      AN    "M 30.0";
      A     "M 0.3";
      JCN   R900;
      JU    E900;

R900: L     L#0;
      T     "DB UTILITY".T90_ET;
      R     "DB UTILITY".T90_DN;

E900: NOP   0;
NETWORK
TITLE =Soft Timer 90 Add Conveyor 4 - Encoder has Stop H - Timer  500mS

      AN    "E 6.6";
      AN    "M 30.0";
      A     "M 0.3";
      AN    "DB UTILITY".Freeze_Sequence_2;
      AN    "DB UTILITY".T90_DN;
      JCN   E901;

      L     "DB UTILITY".T90_ET;
      L     "DB UTILITY".Scan_Cycle_Previous;
      ITD   ;
      +D    ;
      T     "DB UTILITY".T90_ET;

E901: NOP   0;
NETWORK
TITLE =Soft Timer 90 Done 500mS

      L     "DB UTILITY".T90_ET;
      L     L#500;
      >=D   ;
      =     "DB UTILITY".T90_DN;
NETWORK
TITLE =Soft Timer 91 Reset

      A     "E 6.6";
      AN    "M 30.0";
      A     "M 0.3";
      JCN   R910;
      JU    E910;

R910: L     L#0;
      T     "DB UTILITY".T91_ET;
      R     "DB UTILITY".T91_DN;

E910: NOP   0;
NETWORK
TITLE =Soft Timer 91 Add

      A     "E 6.6";
      AN    "M 30.0";
      A     "M 0.3";
      AN    "DB UTILITY".Freeze_Sequence_2;
      AN    "DB UTILITY".T91_DN;
      JCN   E911;

      L     "DB UTILITY".T91_ET;
      L     "DB UTILITY".Scan_Cycle_Previous;
      ITD   ;
      +D    ;
      T     "DB UTILITY".T91_ET;

E911: NOP   0;
NETWORK
TITLE =Soft Timer 91 Done 500mS
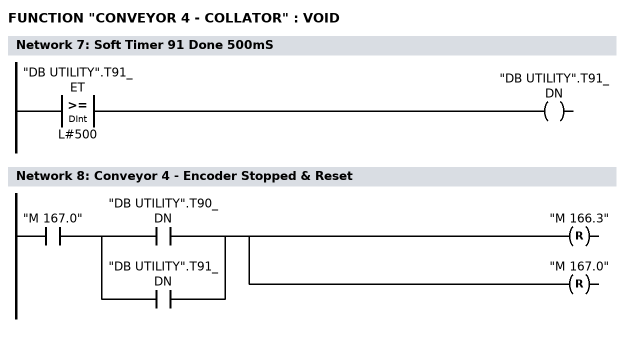

      L     "DB UTILITY".T91_ET;
      L     L#500;
      >=D   ;
      =     "DB UTILITY".T91_DN;
NETWORK
TITLE =Conveyor 4 - Encoder Stopped & Reset

      A     "M 167.0";
      A(    ;
      O     "DB UTILITY".T90_DN;
      O     "DB UTILITY".T91_DN;
      )     ;
      R     "M 166.3";
      R     "M 167.0";
NETWORK
TITLE =Conveyor 4 - Packet Length - Measurements

      A     "B 6.7";
      A     "M 31.1";
      S     "M 166.2"; // Counter 2 Gate - Set
      =     #COUNTER_TRIGGER;
//;
      A     "M 166.2"; // Counter 2
      =     "FM350 DB".CONTROL_SIGNALS.SW_GATE2; // C4 Length Count
//;
      A     "M 166.2"; // Counter 2
      O     "B 6.4";
      FP    "FP 149.4";
      JNB   NRAZ;
      L     0; // Reset First
      T     "COLLATORS DB".Packet_Length_C4_mS;

NRAZ: A     "M 166.2"; // Counter 2
      JNB   NCNT;
      L     "COLLATORS DB".Packet_Length_C4_mS;
      L     "DB UTILITY".Scan_Cycle_Previous;
      +I    ;
      T     "COLLATORS DB".Packet_Length_C4_mS; // Added ScanCycles

NCNT: A     "M 166.2"; // Counter 2
      AN    "B 6.4";
      AN    "B 6.7";
      JNB   B067;
      L     "FM350 DB".ACT_CNTV2; // C4 Length Count
      T     "COLLATORS DB".PacketLength_C4; // Encoder Pulses - Length
      T     #PACKET_LENGTH_4;
//;
      L     #PACKET_LENGTH_4;
      ITD   ;
      DTR   ;
      L     2.000000e-01;
      *R    ;
      RND   ;


      T     "COLLATORS DB".Frac_Packet_Length_C4;


      L     #PACKET_LENGTH_4;
      +I    ;
      T     "COLLATORS DB".Packet_Length_Frac_C4;
      R     "M 166.2"; // Counter 2 Gate - Reset
      S     "M 167.1";
      S     "M 167.4";

B067: NOP   0;














NETWORK
TITLE =Packet Length Measurements [mm] - While Collating

//    A     "HOUSE_KEEPING DB".C4_First_Collating
      A     "B 6.7"; // C4 InFeed Sens - New Packet
      FP    "FP 226.1";
      A     "A 44.3";
      JCN   NPRT;

      L     "FM350 DB".ACT_CNTV3;
      T     "HOUSE_KEEPING DB".C4_Encoder_READ_Mem;

//NPRT: A     "HOUSE_KEEPING DB".C4_First_Collating
NPRT: AN    "B 6.7"; // C4 InFeed Sens - New Packet End
      FP    "FP 226.2";
      JCN   NTKE;

      L     "FM350 DB".ACT_CNTV3;
      L     "HOUSE_KEEPING DB".C4_Encoder_READ_Mem;
      -I    ;
      T     "HOUSE_KEEPING DB".C4_Packet_Length_ep; // C4 Packet Length [ep]
      DTR   ;
//;
      L     6.350000e+00; //  Encoder Wheel 635mm / 100 PPR  [mm/pulse]
      *R    ;
      RND   ;
      T     "HOUSE_KEEPING DB".C4_Packet_Length_mm;

NTKE: NOP   0;
NETWORK
TITLE =Packet Length Measurements [mS] - While Transfering to C5

      A     "M 31.6"; // C4 Transfer Step
      A     "B 7.0"; // C4 This Packet Exiting
      JCN   NMSR;
      L     "HOUSE_KEEPING DB".C4_Added_Scans_mS;
      L     "DB UTILITY".Scan_Cycle_Previous;
      +I    ;
      T     "HOUSE_KEEPING DB".C4_Added_Scans_mS; // Adding mS

NMSR: A     "M 31.6"; // C4 Transfer Step
      AN    "B 7.0"; // C4 This Packet Exiting Done
      FP    "FP 226.3";
      JCN   NLNT;

      L     "HOUSE_KEEPING DB".C4_Added_Scans_mS;
      T     "HOUSE_KEEPING DB".C4_Packet_Length_mS; // Packet Length mS @ 31 m/min
//;
      L     0;
      T     "HOUSE_KEEPING DB".C4_Added_Scans_mS; // Packet Length mS - Zeroed

NLNT: NOP   0;
NETWORK
TITLE =Between Packets Spaces - Measurements [mm]
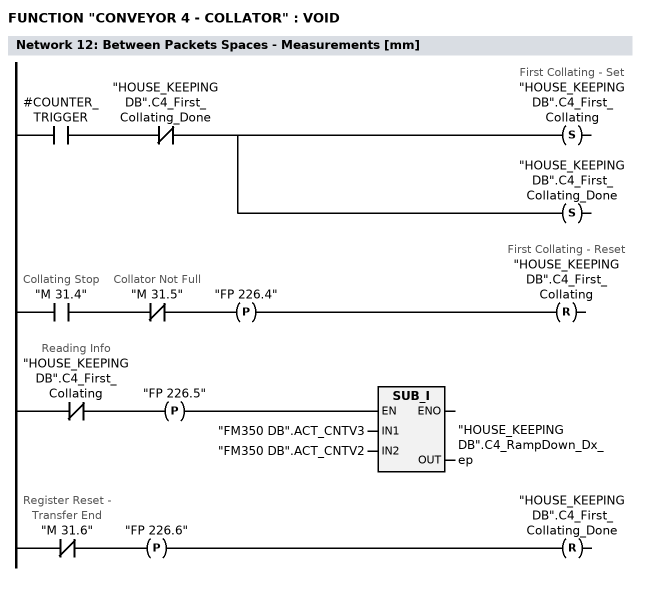

      A     #COUNTER_TRIGGER;
      AN    "HOUSE_KEEPING DB".C4_First_Collating_Done;
      S     "HOUSE_KEEPING DB".C4_First_Collating; // First Collating - Set
      S     "HOUSE_KEEPING DB".C4_First_Collating_Done;
//;
      A     "M 31.4"; // Collating Stop
      AN    "M 31.5"; // Collator Not Full
      FP    "FP 226.4";
      R     "HOUSE_KEEPING DB".C4_First_Collating; // First Collating - Reset
//;
      AN    "HOUSE_KEEPING DB".C4_First_Collating; // Reading Info
      FP    "FP 226.5";
      JCN   N1ST;

      L     "FM350 DB".ACT_CNTV3;
      L     "FM350 DB".ACT_CNTV2;
      -I    ;
      T     "HOUSE_KEEPING DB".C4_RampDown_Dx_ep;

N1ST: NOP   0;

      AN    "M 31.6"; // Register Reset - Transfer End
      FP    "FP 226.6";
      R     "HOUSE_KEEPING DB".C4_First_Collating_Done;
NETWORK
TITLE =Conveyor 4 - Surface Length Left (PulseUnit) - Measurements

      A     "M 31.1";
      S     "M 166.3";
//;
      A     "M 166.3";
      AN    "M 31.7";
      =     "FM350 DB".CONTROL_SIGNALS.SW_GATE3;
//;
      A     "M 166.3";
      A     "M 31.1";
      JNB   M663;
      L     "COLLATORS DB".Surface_Length_C4;
      L     "FM350 DB".ACT_CNTV3;
      -D    ;
      T     "COLLATORS DB".Surface_Left_C4;
      L     0;
      >=I   ;
      JNB   T004;
      L     "COLLATORS DB".Surface_Left_C4;
      T     "COLLATORS DB".Surface_Length_Left_C4;

T004: CLR   ;

M663: CLR   ;
NETWORK
TITLE =Conveyor 4 - Space Between - Calculator

      A     "M 167.1";
      FP    "FP 154.2";
      JNB   M581;
      L     "COLLATORS DB".Surface_Left_C4;
      L     "COLLATORS DB".Frac_Packet_Length_C4;
      -I    ;
      T     "MW 214";

M581: CLR   ;

      A     "M 167.1";
      JNB   M671;
      A(    ;
      L     "COLLATORS DB".Surface_Left_C4;
      L     "MW 214";
      <=I   ;
      )     ;
      R     "M 167.1";

M671: CLR   ;
NETWORK
TITLE =Conveyor 4 - Collating Length Manager

      A     "M 166.3";
      AN    "M 30.4";
      A     "M 31.4";
      JNB   M304;
      L     "COLLATORS DB".Surface_Left_C4;
      L     "COLLATORS DB".Packet_Length_Frac_C4;
      <I    ;
      S     "M 30.4";

M304: CLR   ;

      A     "M 10.1";
      FP    "FP 154.7";
      O     "M 31.7";
      R     "M 30.4";
NETWORK
TITLE =Packet Length to HMI + Hysteresis

      A     "M 167.4";
      JNB   C167;
      A(    ;
      A(    ;
      L     "MW 202";
      L     "MW 204";
      >I    ;
      )     ;
      O     ;
      A(    ;
      L     "MW 202";
      L     "MW 206";
      <I    ;
      )     ;
      )     ;
      JNB   BYP5;
      L     "MW 202";
      T     "HMI_DB".WORD_PACKET_LENGTH;

BYP5: CLR   ;

      L     "MW 202";
      L     3.000000e+00;
      *R    ;
      L     1.000000e+02;
      /R    ;
      T     #R_TUBE_PERCENT;
      TRUNC ;
//     T     "COLLATORS DB".Ecoder_Wheel_Circ_C4
      T     #W_TUBE_PERCENT;
//;
      L     #W_TUBE_PERCENT;
      L     "MW 202";
      +I    ;
      T     "MW 204";
//;
      L     #W_TUBE_PERCENT;
      L     "MW 202";
      -I    ;
      T     "MW 206";
//;
      CLR   ;
      =     "M 167.4";

C167: CLR   ;
NETWORK
TITLE =Collator
//Collator House Keeping


NETWORK
TITLE =Collator Conveyor 4 - Clearing
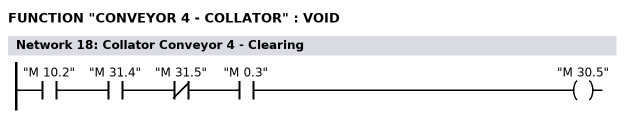

      A     "M 10.2";
      A     "M 31.4";
      AN    "M 31.5";
      A     "M 0.3";
      =     "M 30.5";
NETWORK
TITLE =Soft Timer 33 Reset - Clearing TimeOut 20s + Freeze Option

      A     "M 30.5";
      A     "A 44.3";
      A     "M 0.3";
      JCN   R331;
      JU    E331;

R331: L     L#0;
      T     "DB UTILITY".T33_ET;
      R     "DB UTILITY".T33_DN;

E331: NOP   0;
NETWORK
TITLE =Soft Timer 33 Add

      A     "M 30.5";
      A     "A 44.3";
      A     "M 0.3";
      AN    "DB UTILITY".Freeze_Sequence_2;
      AN    "DB UTILITY".T33_DN;
      JCN   E332;

      L     "DB UTILITY".T33_ET;
      L     "DB UTILITY".Scan_Cycle_Previous;
      ITD   ;
      +D    ;
      T     "DB UTILITY".T33_ET;

E332: NOP   0;
NETWORK
TITLE =Soft Timer 33 Done 20s

      L     "DB UTILITY".T33_ET;
      L     L#20000;
      >=D   ;
      =     "DB UTILITY".T33_DN;
NETWORK
TITLE =Collator Conveyor 4 - Clearing Surface - Run 2K Encoder Counts

      A     "M 30.5";
      A     "A 44.3";
      A     "M 0.3";
      JNB   M305;
      A(    ;
      L     "FM350 DB".ACT_CNTV2;
      L     2000;
      >I    ;
      )     ;
      =     "M 30.3";

M305: CLR   ;
NETWORK
TITLE =Collator Conveyor 4 - Packet at the End !
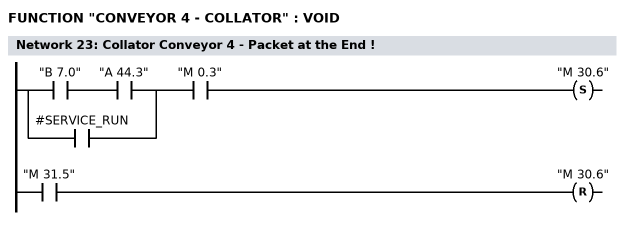

      A     "B 7.0";
      A     "A 44.3";
      O     #SERVICE_RUN;
      A     "M 0.3";
      S     "M 30.6";
//;
      A     "M 31.5";
      R     "M 30.6";
NETWORK
TITLE =Soft Timer 31 Reset - InFeed TimeOut 5s With Freeze Option

      A     "M 31.2";
      AN    "M 31.4";
      A     "A 44.3";
      A     "M 0.3";
      JCN   R311;
      JU    E311;

R311: L     L#0;
      T     "DB UTILITY".T31_ET;
      R     "DB UTILITY".T31_DN;

E311: NOP   0;
NETWORK
TITLE =Soft Timer 31 Add

      A     "M 31.2";
      AN    "M 31.4";
      A     "A 44.3";
      A     "M 0.3";
      AN    "DB UTILITY".Freeze_Sequence_2;
      AN    "DB UTILITY".T31_DN;
      JCN   E312;

      L     "DB UTILITY".T31_ET;
      L     "DB UTILITY".Scan_Cycle_Previous;
      ITD   ;
      +D    ;
      T     "DB UTILITY".T31_ET;

E312: NOP   0;
NETWORK
TITLE =Soft Timer 31 Done 5s
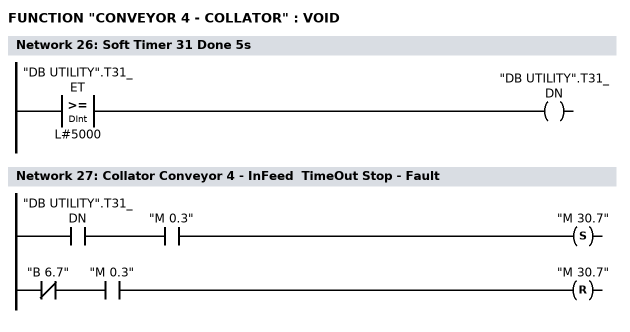

      L     "DB UTILITY".T31_ET;
      L     L#5000;
      >=D   ;
      =     "DB UTILITY".T31_DN;
NETWORK
TITLE =Collator Conveyor 4 - InFeed  TimeOut Stop - Fault

      A     "DB UTILITY".T31_DN;
      A     "M 0.3";
      S     "M 30.7";
//;
      AN    "B 6.7";
      A     "M 0.3";
      R     "M 30.7";
NETWORK
TITLE =Collator
//Collator Steps


NETWORK
TITLE =Collator Conveyor 4 - Steps Register - Reset

      A(    ;
      O     "M 31.7";
      O     "DB UTILITY".T33_DN;
      O     #INITIALISATION;
      O     "DB UTILITY".Conveyor_4_Disable;
      )     ;
      A     "M 0.3";
      JNB   INIT;
      L     W#16#0;
      T     "MW 31";
      S     "M 167.0";

INIT: CLR   ;
NETWORK
TITLE =Step 5N1  - Power ON
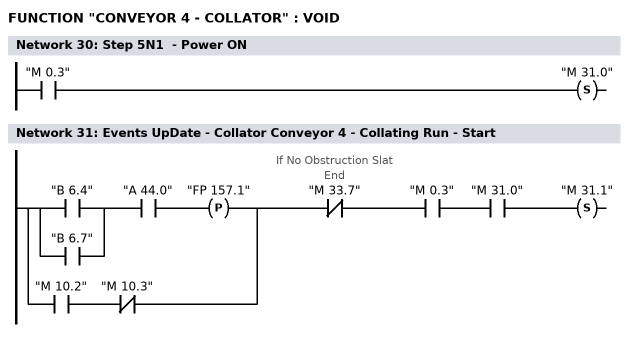

      A     "M 0.3";
      S     "M 31.0";
NETWORK
TITLE =Events UpDate - Collator Conveyor 4 - Collating Run - Start

      A(    ;
      A(    ;
      O     "B 6.4";
      O     "B 6.7";
      )     ;
      A     "A 44.0";
      FP    "FP 157.1";
      O     ;
      A     "M 10.2";
      AN    "M 10.3";
      )     ;
      AN    "M 33.7"; // If No Obstruction Slat End
      A     "M 0.3";
      A     "M 31.0";
      S     "M 31.1";
NETWORK
TITLE =Soft Timer 29 Reset - LB Obstruction Alarm 10s + Freeze Option

      A(    ;
      O     "B 6.4";
      O     "B 6.7";
      )     ;
      AN    "A 44.0";
      JCN   R281;
      JU    E281;

R281: L     L#0;
      T     "DB UTILITY".T29_ET;
      R     "DB UTILITY".T29_DN;

E281: NOP   0;
NETWORK
TITLE =Soft Timer 29 Add

      A(    ;
      O     "B 6.4";
      O     "B 6.7";
      )     ;
      AN    "A 44.0";
      AN    "DB UTILITY".Freeze_Sequence_2;
      AN    "DB UTILITY".T29_DN;
      JCN   E282;

      L     "DB UTILITY".T29_ET;
      L     "DB UTILITY".Scan_Cycle_Previous;
      ITD   ;
      +D    ;
      T     "DB UTILITY".T29_ET;

E282: NOP   0;
NETWORK
TITLE =Soft Timer 29 Done 10s
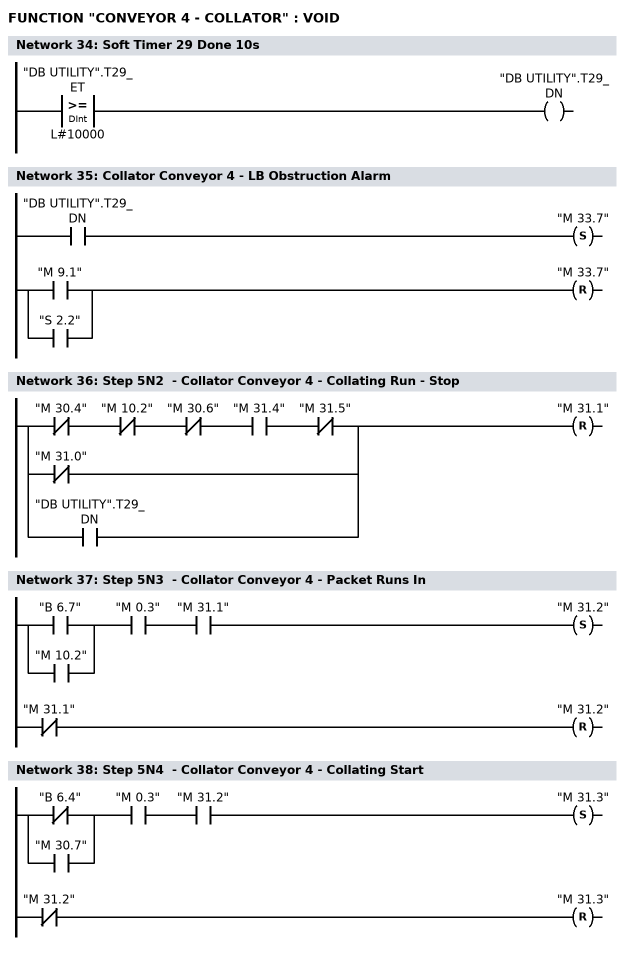

      L     "DB UTILITY".T29_ET;
      L     L#10000;
      >=D   ;
      =     "DB UTILITY".T29_DN;
NETWORK
TITLE =Collator Conveyor 4 - LB Obstruction Alarm

      A     "DB UTILITY".T29_DN;
      S     "M 33.7";
//;
      A(    ;
      O     "M 9.1";
      O     "S 2.2";
      )     ;
      R     "M 33.7";
NETWORK
TITLE =Step 5N2  - Collator Conveyor 4 - Collating Run - Stop

      A(    ;
      AN    "M 30.4";
      AN    "M 10.2";
      AN    "M 30.6";
      A     "M 31.4";
      AN    "M 31.5";
      ON    "M 31.0";
      O     "DB UTILITY".T29_DN;
      )     ;
      R     "M 31.1";
NETWORK
TITLE =Step 5N3  - Collator Conveyor 4 - Packet Runs In

      A(    ;
      O     "B 6.7";
      O     "M 10.2";
      )     ;
      A     "M 0.3";
      A     "M 31.1";
      S     "M 31.2";
//;
      AN    "M 31.1";
      R     "M 31.2";
NETWORK
TITLE =Step 5N4  - Collator Conveyor 4 - Collating Start

      A(    ;
      ON    "B 6.4";
      O     "M 30.7";
      )     ;
      A     "M 0.3";
      A     "M 31.2";
      S     "M 31.3";
//;
      AN    "M 31.2";
      R     "M 31.3";
NETWORK
TITLE =Step 5N5  - Collator Conveyor 4 - Collating Stop

      A(    ;
      AN    "B 6.7";
      AN(   ;
      AN    "M 10.2";
      A     "M 167.1";
      )     ;
      O     "M 30.7";
      )     ;
      A     "M 0.3";
      A     "M 31.3";
      S     "M 31.4";
//;
      AN    "M 31.3";
      R     "M 31.4";
NETWORK
TITLE =Step 5N6  - Collator Conveyor 4 - Full - Start Transfer
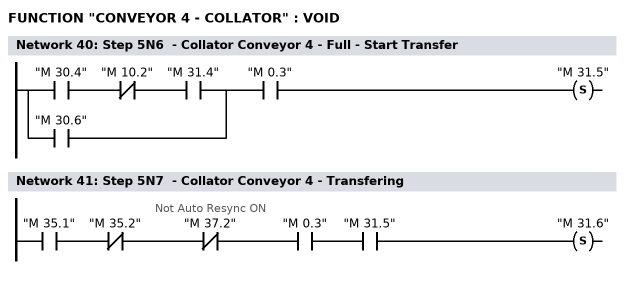

      A(    ;
      A     "M 30.4";
      AN    "M 10.2";
      A     "M 31.4";
      O     "M 30.6";
      )     ;
      A     "M 0.3";
      S     "M 31.5";
NETWORK
TITLE =Step 5N7  - Collator Conveyor 4 - Transfering

      A     "M 35.1";
      AN    "M 35.2";
      AN    "M 37.2"; // Not Auto Resync ON
      A     "M 0.3";
      A     "M 31.5";
      S     "M 31.6";
NETWORK
TITLE =Soft Timer 32 Reset - Transfer TimeOut 20s + Freeze Option

      A     "M 31.6";
      AN    "M 31.7";
      A     "A 44.3";
      A     "M 0.3";
      JCN   R321;
      JU    E321;

R321: L     L#0;
      T     "DB UTILITY".T32_ET;
      R     "DB UTILITY".T32_DN;

E321: NOP   0;
NETWORK
TITLE =Soft Timer 32 Add

      A     "M 31.6";
      AN    "M 31.7";
      A     "A 44.3";
      A     "M 0.3";
      AN    "DB UTILITY".Freeze_Sequence_2;
      AN    "DB UTILITY".T32_DN;
      JCN   E322;

      L     "DB UTILITY".T32_ET;
      L     "DB UTILITY".Scan_Cycle_Previous;
      ITD   ;
      +D    ;
      T     "DB UTILITY".T32_ET;

E322: NOP   0;
NETWORK
TITLE =Soft Timer 32 Done 20s
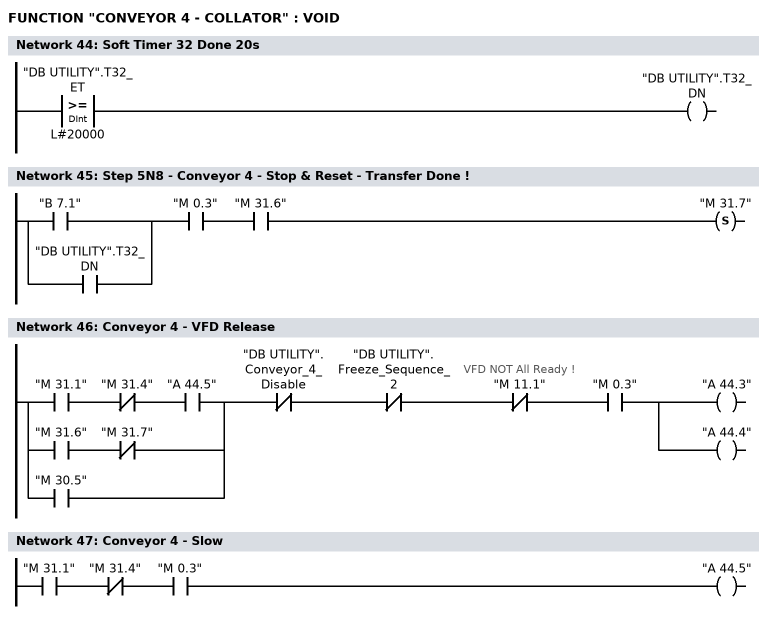

      L     "DB UTILITY".T32_ET;
      L     L#20000;
      >=D   ;
      =     "DB UTILITY".T32_DN;
NETWORK
TITLE =Step 5N8 - Conveyor 4 - Stop & Reset - Transfer Done !

      A(    ;
      O     "B 7.1";
      O     "DB UTILITY".T32_DN;
      )     ;
      A     "M 0.3";
      A     "M 31.6";
      S     "M 31.7";
NETWORK
TITLE =Conveyor 4 - VFD Release

      A(    ;
      A     "M 31.1";
      AN    "M 31.4";
      A     "A 44.5";
      O     ;
      A     "M 31.6";
      AN    "M 31.7";
      O     "M 30.5";
      )     ;
      AN    "DB UTILITY".Conveyor_4_Disable;
      AN    "DB UTILITY".Freeze_Sequence_2;
      AN    "M 11.1"; // VFD NOT All Ready !
      A     "M 0.3";
      =     "A 44.3";
      =     "A 44.4";
NETWORK
TITLE =Conveyor 4 - Slow

      A     "M 31.1";
      AN    "M 31.4";
      A     "M 0.3";
      =     "A 44.5";
END_FUNCTION

FUNCTION "CONVEYOR 5 - LINK" : VOID
TITLE =Conveyor 5 - Link   Pos.7
//Using "Soft Timer" cause S5T Timer cannot Pause/Freeze !...
NAME : POS_7
VERSION : 0.0


VAR_TEMP
  MAIN_SERVICE_2_SW : BOOL ;
  SERVICE_RUN : BOOL ;
  INITIALISATION : BOOL ;
END_VAR
BEGIN
NETWORK
TITLE =Conveyor 5 - Service

      A     "HMI_DB".ALL_SERVICE_ENABLE_SW;
      A     "HMI_DB".CONVEYOR_5_SERVICE_SW;
      A     "HMI_DB".SERVICE_SW_2_STATUS;
      =     #MAIN_SERVICE_2_SW;
//;
      A     #MAIN_SERVICE_2_SW;
      O     "M 34.1";
      JNB   CON5;
//;
      A     "HMI_DB".HMI_CONVEYOR_5_TEST_SSW;
      AN    "A 44.3";
      =     #SERVICE_RUN;
      S     "DB UTILITY".Conveyor_4_Disable;
//;
      A     "HMI_DB".SERVICE_INIT_PB;
      =     #INITIALISATION;
//;
      AN    #MAIN_SERVICE_2_SW;
      R     "HMI_DB".HMI_CONVEYOR_5_TEST_SSW;
      R     "DB UTILITY".Conveyor_4_Disable;

CON5: R     #SERVICE_RUN;
      R     #INITIALISATION;
      FP    "FP 158.5";
      =     "M 34.1";

NETWORK
TITLE =Service Mode
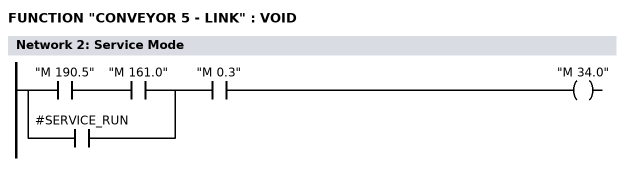

      A(    ;
      A     "M 190.5";
      A     "M 161.0";
      O     ;
      A     #SERVICE_RUN;
      )     ;
      A     "M 0.3";
      =     "M 34.0";

NETWORK
TITLE =Conveyor 5 - Steps Register - Reset

      A(    ;
      A     "M 35.1";
      AN    "M 35.2";
      A     "DB UTILITY".T35_DN;
      O     "M 35.4";
      O     #INITIALISATION;
      O     "DB UTILITY".Conveyor_5_Disable;
      )     ;
      A     "M 0.3";
      JC    M001;
      JU    M002;

M001: L     W#16#0;
      T     "MW 35";
      T     "HMI DB NEW".CONV_5_COUNT;

M002: NOP   0;

NETWORK
TITLE =Step 6N1 - Power ON
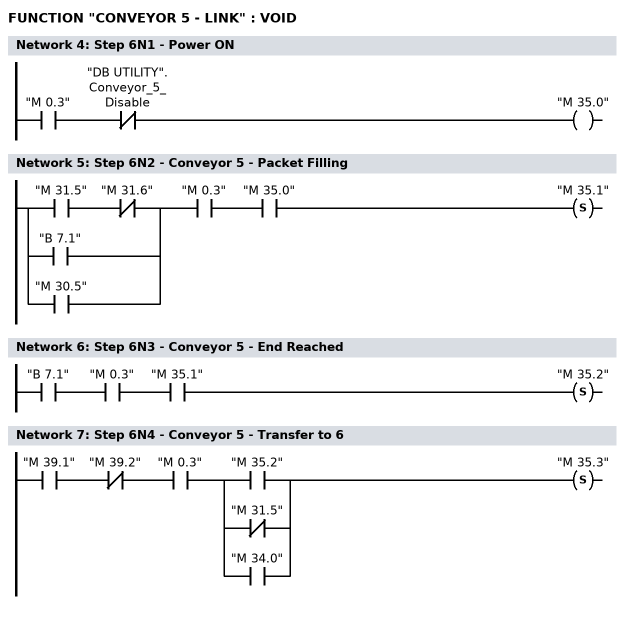

      A     "M 0.3";
      AN    "DB UTILITY".Conveyor_5_Disable;
      =     "M 35.0";

NETWORK
TITLE =Step 6N2 - Conveyor 5 - Packet Filling

      A(    ;
      A     "M 31.5";
      AN    "M 31.6";
      O     "B 7.1";
      O     "M 30.5";
      )     ;
      A     "M 0.3";
      A     "M 35.0";
      S     "M 35.1";

NETWORK
TITLE =Step 6N3 - Conveyor 5 - End Reached

      A     "B 7.1";
      A     "M 0.3";
      A     "M 35.1";
      S     "M 35.2";

NETWORK
TITLE =Step 6N4 - Conveyor 5 - Transfer to 6

      A     "M 39.1";
      AN    "M 39.2";
      A     "M 0.3";
      A(    ;
      O     "M 35.2";
      ON    "M 31.5";
      O     "M 34.0";
      )     ;
      S     "M 35.3";

NETWORK
TITLE =Soft Timer 35 Reset

      A(    ;
      A     "M 35.1";
      AN    "M 35.2";
      O     ;
      A     "M 35.3";
      AN    "M 35.4";
      A     "A 45.0";
      )     ;
      A     "M 0.3";
      JCN   R351;
      JU    E351;

R351: L     L#0;
      T     "DB UTILITY".T35_ET;
      R     "DB UTILITY".T35_DN;

E351: NOP   0;

NETWORK
TITLE =Soft Timer 35 Add

      A(    ;
      A     "M 35.1";
      AN    "M 35.2";
      O     ;
      A     "M 35.3";
      AN    "M 35.4";
      A     "A 45.0";
      )     ;
      A     "M 0.3";
      JCN   E352;
//;
      A     "DB UTILITY".Freeze_Sequence_2;
      A     "M 35.1";
      AN    "M 35.2";
      JC    E352;
//;
      AN    "DB UTILITY".T35_DN;
      JCN   E352;
//;
      L     "DB UTILITY".T35_ET;
      L     "DB UTILITY".Scan_Cycle_Previous;
      ITD   ;
      +D    ;
      T     "DB UTILITY".T35_ET;

E352: NOP   0;

NETWORK
TITLE =Soft Timer 35 Done 30s

      L     "DB UTILITY".T35_ET;
      L     L#30000; // [mS]
      >=D   ;
      =     "DB UTILITY".T35_DN;

NETWORK
TITLE =Automatic Re-Synchronization
//In Order to keep Synchronized,
//if Every Conditions are there, Conveyor 5 will do a Synchro Run 13sec after
//every 5 runs !
      A     "A 45.0"; // Count runs
      FP    "FP 169.7";
      JNB   ARS1;

      L     "MW 220"; // Count up
      L     1;
      +I    ;
      T     "MW 220";
//;
      L     10;
      >=I   ;
      JNB   ARS1;
//;
      S     "M 37.3"; // ARM after 5 runs
      L     0;
      T     "MW 220";

ARS1: NOP   0;

      A     "M 37.3"; // ARMED
      AN    "M 37.2"; // NOT already running
      AN    "DB UTILITY".Freeze_Sequence_2;
      AN    "A 45.0"; // wait end of run
      A     "M 35.0"; // power ON
      AN    "M 35.4"; // not in reset/stop
      JNB   ARS2;
//;
      L     "HMI_DB".CONV_4_COUNT; // Conveyor 4 Must be <= 2
      L     3;
      <I    ;
      JNB   ARS2;
//;
      L     "HMI_DB".CONV_5_COUNT;
      L     0; // Conveyor 5 Must NOT be Empty
      >I    ;
      JNB   ARS2;
//;
      L     "HMI_DB".CONV_6_COUNT;
      L     0; // Conveyor 6 Must be Empty
      ==I   ;
      JNB   ARS2;
//;
      AN    "B 7.2"; // Conveyor 6 Must be Empty
      AN    "M 10.0"; // Not Clearing
      JNB   ARS2;
//;
      S     "M 37.2"; // START 13s RUN
      R     "M 37.3"; // DISARM

ARS2: NOP   0;

      A     "M 37.2"; // Re-Sync ON
      L     S5T#13S;
      SD    "Timer 64";
//;
      A     "Timer 64"; // End Re-Sync if TimeOut 13s
      O     "B 7.1"; // or if Packet at END Sensor
      R     "M 37.2"; // Re-Sync OFF
NETWORK
TITLE =Automatic Re-Synchronization - Arm Timeout
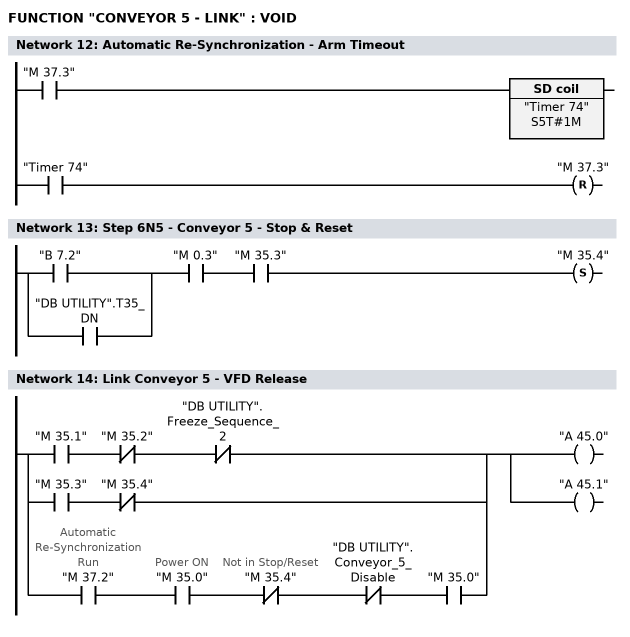

      A     "M 37.3";
      L     S5T#1M;
      SD    "Timer 74";
//;
      A     "Timer 74";
      R     "M 37.3";
NETWORK
TITLE =Step 6N5 - Conveyor 5 - Stop & Reset

      A(    ;
      O     "B 7.2";
      O     "DB UTILITY".T35_DN;
      )     ;
      A     "M 0.3";
      A     "M 35.3";
      S     "M 35.4";

NETWORK
TITLE =Link Conveyor 5 - VFD Release


      A(    ;
      A(    ;
      A     "M 35.1";
      AN    "M 35.2";
      AN    "DB UTILITY".Freeze_Sequence_2;
      )     ;
      O     ;
      A     "M 35.3";
      AN    "M 35.4";
      )     ;
      O     ;
      A(    ;
      A     "M 37.2"; // Automatic Re-Synchronization Run
      A     "M 35.0"; // Power ON
      AN    "M 35.4"; // Not in Stop/Reset
      )     ;
      AN    "DB UTILITY".Conveyor_5_Disable;
      A     "M 35.0";
      =     "A 45.0";
      =     "A 45.1";
END_FUNCTION

FUNCTION "CONVEYOR 6 - FLIP DELIV." : VOID
TITLE =Conveyor 6 - Delivery to Flipper Pos.8
//
NAME : POS_8
VERSION : 0.0


VAR_TEMP
  MAIN_SERVICE_2_SW : BOOL ;
  SERVICE_RUN : BOOL ;
  INITIALISATION : BOOL ;
END_VAR
BEGIN
NETWORK
TITLE =Slat Conveyor - Service

      A     "HMI_DB".ALL_SERVICE_ENABLE_SW;
      A     "HMI_DB".CONVEYOR_6_SERVICE_SW;
      A     "HMI_DB".SERVICE_SW_2_STATUS;
      =     #MAIN_SERVICE_2_SW;
//;
      A     #MAIN_SERVICE_2_SW;
      O     "M 38.1";
      JNB   CON6;
      A     "HMI_DB".HMI_CONVEYOR_6_TEST_SSW;
      =     #SERVICE_RUN;
      S     "DB UTILITY".Conveyor_5_Disable;
//;
      AN    #MAIN_SERVICE_2_SW;
      R     "HMI_DB".HMI_CONVEYOR_6_TEST_SSW;
      R     "DB UTILITY".Conveyor_5_Disable;

CON6: R     #SERVICE_RUN;
      R     #INITIALISATION;
      FP    "FP 158.6";
      =     "M 38.1";
NETWORK
TITLE =Flipper Delivery Conveyor 6 - Running TimeOut  30s
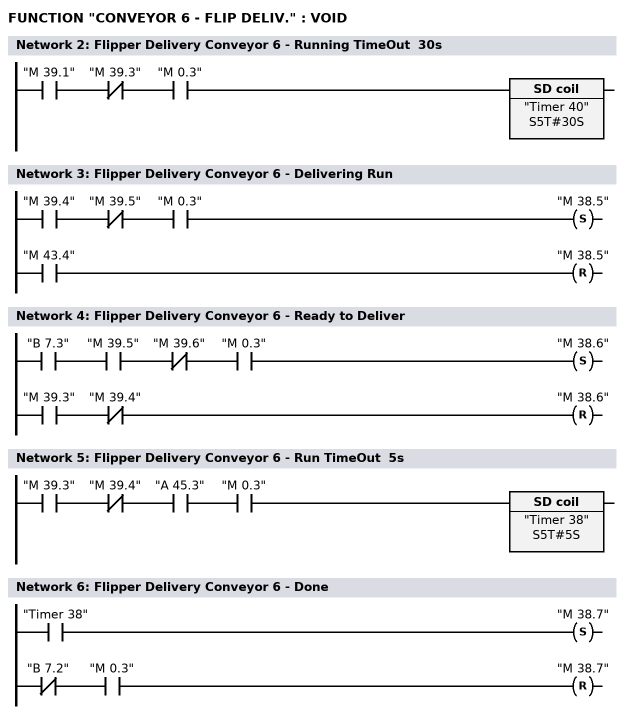

      A     "M 39.1";
      AN    "M 39.3";
      A     "M 0.3";
      L     S5T#30S;
      SD    "Timer 40";
NETWORK
TITLE =Flipper Delivery Conveyor 6 - Delivering Run

      A     "M 39.4";
      AN    "M 39.5";
      A     "M 0.3";
      S     "M 38.5";
//;
      A     "M 43.4";
      R     "M 38.5";
NETWORK
TITLE =Flipper Delivery Conveyor 6 - Ready to Deliver

      A     "B 7.3";
      A     "M 39.5";
      AN    "M 39.6";
      A     "M 0.3";
      S     "M 38.6";
//;
      A     "M 39.3";
      AN    "M 39.4";
      R     "M 38.6";
NETWORK
TITLE =Flipper Delivery Conveyor 6 - Run TimeOut  5s

      A     "M 39.3";
      AN    "M 39.4";
      A     "A 45.3";
      A     "M 0.3";
      L     S5T#5S;
      SD    "Timer 38";
NETWORK
TITLE =Flipper Delivery Conveyor 6 - Done

      A     "Timer 38";
      S     "M 38.7";
//;
      AN    "B 7.2";
      A     "M 0.3";
      R     "M 38.7";
NETWORK
TITLE =Conveyor 6 - Steps Register - Reset

      A(    ;
      O     "M 39.6";
      O     "Timer 40";
      O     #INITIALISATION;
      O     "DB UTILITY".Conveyor_6_Disable;
      )     ;
      A     "M 0.3";
      JC    M001;
      JU    M002;

M001: L     W#16#0;
      T     "MW 39";
      T     "MB 41";
      T     "HMI DB NEW".CONV_6_COUNT;

M002: NOP   0;
NETWORK
TITLE =Step 7N1 - Power ON
